Fanuc KAREL source: kt00089.KL

-- PROVISIONAL review KL for V770-1; original PC SHA256 ca172fed33100f4c6590c7e8202e99a3473a7f78a9453ade4241603317150010
-- Incomplete behavior may be omitted. Consult companion uncertainty JSON. Do not deploy.
PROGRAM KT00089
%NOLOCKGROUP
VAR
  I2 : INTEGER
  OUT : INTEGER
-- UNRESOLVED_DECL H1 type=002017
BEGIN
  -- UNRESOLVED_PC offsets 5-19; opcodes 2E,22,9D,33,B4
  -- UNRESOLVED_PC offsets 24-35; opcodes 2E,23
  -- UNRESOLVED_PC offsets 40-62; opcodes 22,9D,33,B3,21,54,23
  -- UNRESOLVED_PC offsets 67-71; opcodes 7F
END KT00089
